//------------------------------------------------------------------------------
// SCADA FUXA : holding registers (FUXA 400001...), REAL = low word first (Float32MLE)
//------------------------------------------------------------------------------
	//--- DIP1500_1
	GVL_COM.COM_DIP1500_1.SCADA_INPUT_MOTOR_SPEED.Word_value[0]                                := GVL_MODBUS.Holding_register_TCP_HMI[0];    // 1 | DIP1500 Motor Speed (low word)
	GVL_COM.COM_DIP1500_1.SCADA_INPUT_MOTOR_SPEED.Word_value[1]                                := GVL_MODBUS.Holding_register_TCP_HMI[1];    // 2 | DIP1500 Motor Speed (high word)
	GVL_COM.COM_DIP1500_1.SCADA_INPUT_MAX_MOTOR_SPEED.Word_value[0]                            := GVL_MODBUS.Holding_register_TCP_HMI[2];    // 3 | DIP1500 Max Motor Speed (low word)
	GVL_COM.COM_DIP1500_1.SCADA_INPUT_MAX_MOTOR_SPEED.Word_value[1]                            := GVL_MODBUS.Holding_register_TCP_HMI[3];    // 4 | DIP1500 Max Motor Speed (high word)
	GVL_COM.COM_DIP1500_1.SCADA_INPUT_RUN_TIME_OR_VOLUME_SETPOINT.Word_value[0]                := GVL_MODBUS.Holding_register_TCP_HMI[4];    // 5 | DIP1500 Run Time Or Volume Setpoint (low word)
	GVL_COM.COM_DIP1500_1.SCADA_INPUT_RUN_TIME_OR_VOLUME_SETPOINT.Word_value[1]                := GVL_MODBUS.Holding_register_TCP_HMI[5];    // 6 | DIP1500 Run Time Or Volume Setpoint (high word)
	GVL_COM.COM_DIP1500_1.SCADA_INPUT_FLOW_RATE_OR_SPEED_CALIBRATION_COEFFICIENT.Word_value[0] := GVL_MODBUS.Holding_register_TCP_HMI[6];    // 7 | DIP1500 Flow Rate Or Speed Calibration Coefficient (low word)
	GVL_COM.COM_DIP1500_1.SCADA_INPUT_FLOW_RATE_OR_SPEED_CALIBRATION_COEFFICIENT.Word_value[1] := GVL_MODBUS.Holding_register_TCP_HMI[7];    // 8 | DIP1500 Flow Rate Or Speed Calibration Coefficient (high word)
	GVL_COM.COM_DIP1500_1.SCADA_INPUT_FOOT_SWITCH_INPUT_MODE                                   := GVL_MODBUS.Holding_register_TCP_HMI[8];    // 9 | DIP1500 Foot Switch Input Mode
	GVL_COM.COM_DIP1500_1.SCADA_INPUT_LIQUID_LEVEL_INPUT_MODE                                  := GVL_MODBUS.Holding_register_TCP_HMI[9];    // 10 | DIP1500 Liquid Level Input Mode
	GVL_COM.COM_DIP1500_1.SCADA_INPUT_STATE_OUTPUT_MODE                                        := GVL_MODBUS.Holding_register_TCP_HMI[10];   // 11 | DIP1500 State Output Mode
	GVL_COM.COM_DIP1500_1.SCADA_INPUT_COMMUNICATION_ADDRESS                                    := GVL_MODBUS.Holding_register_TCP_HMI[11];   // 12 | DIP1500 Communication Address
	GVL_COM.COM_DIP1500_1.SCADA_INPUT_BAUD_RATE_INDEX                                          := GVL_MODBUS.Holding_register_TCP_HMI[12];   // 13 | DIP1500 Baud Rate Index


//------------------------------------------------------------------------------
// HMI : coils (1001...)
//------------------------------------------------------------------------------
	//--- DOSENSOR_1
	GVL_COM.COM_DOSENSOR_1.HMI_INPUT_CALIBRATION_HIGH := GVL_MODBUS.Coils_TCP_HMI[125].0;   // 1001 | DO Calibration High
	GVL_COM.COM_DOSENSOR_1.HMI_INPUT_CALIBRATION_LOW  := GVL_MODBUS.Coils_TCP_HMI[125].1;   // 1002 | DO Calibration Low
	GVL_COM.COM_DOSENSOR_1.HMI_INPUT_LOCAL_REQUEST    := GVL_MODBUS.Coils_TCP_HMI[125].7;   // 1008 | DO Sensor Local Request
	GVL_COM.COM_DOSENSOR_1.HMI_INPUT_AUTO_REQUEST     := GVL_MODBUS.Coils_TCP_HMI[126].0;   // 1009 | DO Sensor Auto Request

	//--- DIP1500_1
	GVL_COM.COM_DIP1500_1.HMI_INPUT_MOTOR_START_STOP   := GVL_MODBUS.Coils_TCP_HMI[125].2;   // 1003 | DIP1500 Motor Start Stop
	GVL_COM.COM_DIP1500_1.HMI_INPUT_MOTOR_DIRECTION    := GVL_MODBUS.Coils_TCP_HMI[125].3;   // 1004 | DIP1500 Motor Direction
	GVL_COM.COM_DIP1500_1.HMI_INPUT_FLASH_SAVE         := GVL_MODBUS.Coils_TCP_HMI[125].4;   // 1005 | DIP1500 Flash Save
	GVL_COM.COM_DIP1500_1.HMI_INPUT_OPERATION_MODE     := GVL_MODBUS.Coils_TCP_HMI[125].5;   // 1006 | DIP1500 Operation Mode
	GVL_COM.COM_DIP1500_1.HMI_INPUT_PARAM_WRITE_ENABLE := GVL_MODBUS.Coils_TCP_HMI[125].6;   // 1007 | DIP1500 Parameter Write Enable
	GVL_COM.COM_DIP1500_1.HMI_INPUT_LOCAL_REQUEST      := GVL_MODBUS.Coils_TCP_HMI[126].1;   // 1010 | DIP1500 Local Request
	GVL_COM.COM_DIP1500_1.HMI_INPUT_AUTO_REQUEST       := GVL_MODBUS.Coils_TCP_HMI[126].2;   // 1011 | DIP1500 Auto Request

	//--- ADM100W_1
	GVL_COM.COM_ADM100W_1.HMI_INPUT_LOCAL_REQUEST := GVL_MODBUS.Coils_TCP_HMI[126].3;   // 1012 | ADM100W Local Request
	GVL_COM.COM_ADM100W_1.HMI_INPUT_AUTO_REQUEST  := GVL_MODBUS.Coils_TCP_HMI[126].4;   // 1013 | ADM100W Auto Request

	//--- UPI_LOCAL_HMI
	GVL_COM.COM_UPI_LOCAL_HMI.HMI_INPUT_LOCAL_REQUEST := GVL_MODBUS.Coils_TCP_HMI[126].5;   // 1014 | Global Local HMI Request
	GVL_COM.COM_UPI_LOCAL_HMI.HMI_INPUT_AUTO_REQUEST  := GVL_MODBUS.Coils_TCP_HMI[126].6;   // 1015 | Global Auto HMI Request


//------------------------------------------------------------------------------
// HMI : holding registers (1001...), REAL = low word first
//------------------------------------------------------------------------------
	//--- DIP1500_1
	GVL_COM.COM_DIP1500_1.HMI_INPUT_MOTOR_SPEED.Word_value[0]                                := GVL_MODBUS.Holding_register_TCP_HMI[1000];   // 1001 | DIP1500 Motor Speed (low word)
	GVL_COM.COM_DIP1500_1.HMI_INPUT_MOTOR_SPEED.Word_value[1]                                := GVL_MODBUS.Holding_register_TCP_HMI[1001];   // 1002 | DIP1500 Motor Speed (high word)
	GVL_COM.COM_DIP1500_1.HMI_INPUT_MAX_MOTOR_SPEED.Word_value[0]                            := GVL_MODBUS.Holding_register_TCP_HMI[1002];   // 1003 | DIP1500 Max Motor Speed (low word)
	GVL_COM.COM_DIP1500_1.HMI_INPUT_MAX_MOTOR_SPEED.Word_value[1]                            := GVL_MODBUS.Holding_register_TCP_HMI[1003];   // 1004 | DIP1500 Max Motor Speed (high word)
	GVL_COM.COM_DIP1500_1.HMI_INPUT_RUN_TIME_OR_VOLUME_SETPOINT.Word_value[0]                := GVL_MODBUS.Holding_register_TCP_HMI[1004];   // 1005 | DIP1500 Run Time Or Volume Setpoint (low word)
	GVL_COM.COM_DIP1500_1.HMI_INPUT_RUN_TIME_OR_VOLUME_SETPOINT.Word_value[1]                := GVL_MODBUS.Holding_register_TCP_HMI[1005];   // 1006 | DIP1500 Run Time Or Volume Setpoint (high word)
	GVL_COM.COM_DIP1500_1.HMI_INPUT_FLOW_RATE_OR_SPEED_CALIBRATION_COEFFICIENT.Word_value[0] := GVL_MODBUS.Holding_register_TCP_HMI[1006];   // 1007 | DIP1500 Flow Rate Or Speed Calibration Coefficient (low word)
	GVL_COM.COM_DIP1500_1.HMI_INPUT_FLOW_RATE_OR_SPEED_CALIBRATION_COEFFICIENT.Word_value[1] := GVL_MODBUS.Holding_register_TCP_HMI[1007];   // 1008 | DIP1500 Flow Rate Or Speed Calibration Coefficient (high word)
	GVL_COM.COM_DIP1500_1.HMI_INPUT_FOOT_SWITCH_INPUT_MODE                                   := GVL_MODBUS.Holding_register_TCP_HMI[1008];   // 1009 | DIP1500 Foot Switch Input Mode
	GVL_COM.COM_DIP1500_1.HMI_INPUT_LIQUID_LEVEL_INPUT_MODE                                  := GVL_MODBUS.Holding_register_TCP_HMI[1009];   // 1010 | DIP1500 Liquid Level Input Mode
	GVL_COM.COM_DIP1500_1.HMI_INPUT_STATE_OUTPUT_MODE                                        := GVL_MODBUS.Holding_register_TCP_HMI[1010];   // 1011 | DIP1500 State Output Mode
	GVL_COM.COM_DIP1500_1.HMI_INPUT_COMMUNICATION_ADDRESS                                    := GVL_MODBUS.Holding_register_TCP_HMI[1011];   // 1012 | DIP1500 Communication Address
	GVL_COM.COM_DIP1500_1.HMI_INPUT_BAUD_RATE_INDEX                                          := GVL_MODBUS.Holding_register_TCP_HMI[1012];   // 1013 | DIP1500 Baud Rate Index

GFC_COM_IN := TRUE;

                
END_FUNCTION

FUNCTION GFC_COM_OUT : BOOL

                  
//==============================================================================
// GFC_COM_OUT
// GVL_COM -> Modbus (GVL_MODBUS) : RTU equipment, SCADA FUXA, HMI
// Simple copies only, no conversion (conversions are done in the FBs)
//==============================================================================

//------------------------------------------------------------------------------
// COM : Modbus RTU, to equipment (write triggers are mapped directly in the slave I/O mapping)
//------------------------------------------------------------------------------
	//--- DIP1500_1
	GVL_MODBUS.DIP1500_Coils          := GVL_COM.COM_DIP1500_1.COM_OUTPUT_COILS;       // Coils 0x0001..0x0004
	GVL_MODBUS.DIP1500_Holding_Cmd    := GVL_COM.COM_DIP1500_1.COM_OUTPUT_HR_CMD;      // Holding registers 0x4001..0x4006
	GVL_MODBUS.DIP1500_Holding_Config := GVL_COM.COM_DIP1500_1.COM_OUTPUT_HR_CONFIG;   // Holding registers 0x400B..0x4011


//------------------------------------------------------------------------------
// SCADA FUXA : discrete inputs (FUXA 100001...)
//------------------------------------------------------------------------------
	//--- DOSENSOR_1
	GVL_MODBUS.Discret_input_TCP_HMI[0].0 := GVL_COM.COM_DOSENSOR_1.SCADA_OUTPUT_FAULT;               // 10001 | Do sensor fault
	GVL_MODBUS.Discret_input_TCP_HMI[0].1 := GVL_COM.COM_DOSENSOR_1.SCADA_OUTPUT_CALIBRATION_DONE;    // 10002 | Do sensor calibration done
	GVL_MODBUS.Discret_input_TCP_HMI[1].4 := GVL_COM.COM_DOSENSOR_1.SCADA_OUTPUT_LOCAL_FUXA_ACTIVE;   // 10013 | DO Sensor Local FUXA Active
	GVL_MODBUS.Discret_input_TCP_HMI[1].5 := GVL_COM.COM_DOSENSOR_1.SCADA_OUTPUT_LOCAL_HMI_ACTIVE;    // 10014 | DO Sensor Local HMI Active

	//--- ADM100W_1
	GVL_MODBUS.Discret_input_TCP_HMI[0].2 := GVL_COM.COM_ADM100W_1.SCADA_OUTPUT_ALARM_1_STATUS;      // 10003 | ADM100W Alarm 1 Status
	GVL_MODBUS.Discret_input_TCP_HMI[0].3 := GVL_COM.COM_ADM100W_1.SCADA_OUTPUT_ALARM_2_STATUS;      // 10004 | ADM100W Alarm 2 Status
	GVL_MODBUS.Discret_input_TCP_HMI[0].4 := GVL_COM.COM_ADM100W_1.SCADA_OUTPUT_ALARM_3_STATUS;      // 10005 | ADM100W Alarm 3 Status
	GVL_MODBUS.Discret_input_TCP_HMI[0].5 := GVL_COM.COM_ADM100W_1.SCADA_OUTPUT_ALARM_4_STATUS;      // 10006 | ADM100W Alarm 4 Status
	GVL_MODBUS.Discret_input_TCP_HMI[0].6 := GVL_COM.COM_ADM100W_1.SCADA_OUTPUT_ALARM_5_STATUS;      // 10007 | ADM100W Alarm 5 Status
	GVL_MODBUS.Discret_input_TCP_HMI[0].7 := GVL_COM.COM_ADM100W_1.SCADA_OUTPUT_ALARM_6_STATUS;      // 10008 | ADM100W Alarm 6 Status
	GVL_MODBUS.Discret_input_TCP_HMI[1].0 := GVL_COM.COM_ADM100W_1.SCADA_OUTPUT_ALARM_7_STATUS;      // 10009 | ADM100W Alarm 7 Status
	GVL_MODBUS.Discret_input_TCP_HMI[1].1 := GVL_COM.COM_ADM100W_1.SCADA_OUTPUT_ALARM_8_STATUS;      // 10010 | ADM100W Alarm 8 Status
	GVL_MODBUS.Discret_input_TCP_HMI[1].2 := GVL_COM.COM_ADM100W_1.SCADA_OUTPUT_ALARM_9_STATUS;      // 10011 | ADM100W Alarm 9 Status
	GVL_MODBUS.Discret_input_TCP_HMI[1].3 := GVL_COM.COM_ADM100W_1.SCADA_OUTPUT_ALARM_10_STATUS;     // 10012 | ADM100W Alarm 10 Status
	GVL_MODBUS.Discret_input_TCP_HMI[2].0 := GVL_COM.COM_ADM100W_1.SCADA_OUTPUT_LOCAL_FUXA_ACTIVE;   // 10017 | ADM100W Local FUXA Active
	GVL_MODBUS.Discret_input_TCP_HMI[2].1 := GVL_COM.COM_ADM100W_1.SCADA_OUTPUT_LOCAL_HMI_ACTIVE;    // 10018 | ADM100W Local HMI Active

	//--- DIP1500_1
	GVL_MODBUS.Discret_input_TCP_HMI[1].6 := GVL_COM.COM_DIP1500_1.SCADA_OUTPUT_LOCAL_FUXA_ACTIVE;   // 10015 | DIP1500 Local FUXA Active
	GVL_MODBUS.Discret_input_TCP_HMI[1].7 := GVL_COM.COM_DIP1500_1.SCADA_OUTPUT_LOCAL_HMI_ACTIVE;    // 10016 | DIP1500 Local HMI Active

	//--- UPI_LOCAL_FUXA
	GVL_MODBUS.Discret_input_TCP_HMI[2].2 := GVL_COM.COM_UPI_LOCAL_FUXA.SCADA_OUTPUT_LOCAL_ACTIVE;   // 10019 | Global Local FUXA Active

	//--- UPI_LOCAL_HMI
	GVL_MODBUS.Discret_input_TCP_HMI[2].3 := GVL_COM.COM_UPI_LOCAL_HMI.SCADA_OUTPUT_LOCAL_ACTIVE;   // 10020 | Global Local HMI Active


//------------------------------------------------------------------------------
// SCADA FUXA : input registers (FUXA 300001...), REAL = low word first (Float32MLE)
//------------------------------------------------------------------------------
	//--- ADM100W_1
	GVL_MODBUS.Input_register_TCP_HMI[0]  := GVL_COM.COM_ADM100W_1.SCADA_OUTPUT_FREQUENCY.Word_value[0];                   // 1 | ADM100W Frequency (low word)
	GVL_MODBUS.Input_register_TCP_HMI[1]  := GVL_COM.COM_ADM100W_1.SCADA_OUTPUT_FREQUENCY.Word_value[1];                   // 2 | ADM100W Frequency (high word)
	GVL_MODBUS.Input_register_TCP_HMI[2]  := GVL_COM.COM_ADM100W_1.SCADA_OUTPUT_L1_L2_VOLTAGE.Word_value[0];               // 3 | ADM100W L1-L2 Voltage (low word)
	GVL_MODBUS.Input_register_TCP_HMI[3]  := GVL_COM.COM_ADM100W_1.SCADA_OUTPUT_L1_L2_VOLTAGE.Word_value[1];               // 4 | ADM100W L1-L2 Voltage (high word)
	GVL_MODBUS.Input_register_TCP_HMI[4]  := GVL_COM.COM_ADM100W_1.SCADA_OUTPUT_L1_N_VOLTAGE.Word_value[0];                // 5 | ADM100W L1-N Voltage (low word)
	GVL_MODBUS.Input_register_TCP_HMI[5]  := GVL_COM.COM_ADM100W_1.SCADA_OUTPUT_L1_N_VOLTAGE.Word_value[1];                // 6 | ADM100W L1-N Voltage (high word)
	GVL_MODBUS.Input_register_TCP_HMI[6]  := GVL_COM.COM_ADM100W_1.SCADA_OUTPUT_L1_CURRENT.Word_value[0];                  // 7 | ADM100W L1 Current (low word)
	GVL_MODBUS.Input_register_TCP_HMI[7]  := GVL_COM.COM_ADM100W_1.SCADA_OUTPUT_L1_CURRENT.Word_value[1];                  // 8 | ADM100W L1 Current (high word)
	GVL_MODBUS.Input_register_TCP_HMI[8]  := GVL_COM.COM_ADM100W_1.SCADA_OUTPUT_L1_ACTIVE_POWER.Word_value[0];             // 9 | ADM100W L1 Active Power (low word)
	GVL_MODBUS.Input_register_TCP_HMI[9]  := GVL_COM.COM_ADM100W_1.SCADA_OUTPUT_L1_ACTIVE_POWER.Word_value[1];             // 10 | ADM100W L1 Active Power (high word)
	GVL_MODBUS.Input_register_TCP_HMI[10] := GVL_COM.COM_ADM100W_1.SCADA_OUTPUT_L1_APPARENT_POWER.Word_value[0];           // 11 | ADM100W L1 Apparent Power (low word)
	GVL_MODBUS.Input_register_TCP_HMI[11] := GVL_COM.COM_ADM100W_1.SCADA_OUTPUT_L1_APPARENT_POWER.Word_value[1];           // 12 | ADM100W L1 Apparent Power (high word)
	GVL_MODBUS.Input_register_TCP_HMI[12] := GVL_COM.COM_ADM100W_1.SCADA_OUTPUT_L1_REACTIVE_POWER.Word_value[0];           // 13 | ADM100W L1 Reactive Power (low word)
	GVL_MODBUS.Input_register_TCP_HMI[13] := GVL_COM.COM_ADM100W_1.SCADA_OUTPUT_L1_REACTIVE_POWER.Word_value[1];           // 14 | ADM100W L1 Reactive Power (high word)
	GVL_MODBUS.Input_register_TCP_HMI[14] := GVL_COM.COM_ADM100W_1.SCADA_OUTPUT_L1_CURRENT_PHASE_ANGLE.Word_value[0];      // 15 | ADM100W L1 Current Phase Angle (low word)
	GVL_MODBUS.Input_register_TCP_HMI[15] := GVL_COM.COM_ADM100W_1.SCADA_OUTPUT_L1_CURRENT_PHASE_ANGLE.Word_value[1];      // 16 | ADM100W L1 Current Phase Angle (high word)
	GVL_MODBUS.Input_register_TCP_HMI[16] := GVL_COM.COM_ADM100W_1.SCADA_OUTPUT_L1_POWER_FACTOR.Word_value[0];             // 17 | ADM100W L1 Power Factor (low word)
	GVL_MODBUS.Input_register_TCP_HMI[17] := GVL_COM.COM_ADM100W_1.SCADA_OUTPUT_L1_POWER_FACTOR.Word_value[1];             // 18 | ADM100W L1 Power Factor (high word)
	GVL_MODBUS.Input_register_TCP_HMI[18] := GVL_COM.COM_ADM100W_1.SCADA_OUTPUT_L1_VOLTAGE_THD.Word_value[0];              // 19 | ADM100W L1 Voltage THD (low word)
	GVL_MODBUS.Input_register_TCP_HMI[19] := GVL_COM.COM_ADM100W_1.SCADA_OUTPUT_L1_VOLTAGE_THD.Word_value[1];              // 20 | ADM100W L1 Voltage THD (high word)
	GVL_MODBUS.Input_register_TCP_HMI[20] := GVL_COM.COM_ADM100W_1.SCADA_OUTPUT_L1_CURRENT_THD.Word_value[0];              // 21 | ADM100W L1 Current THD (low word)
	GVL_MODBUS.Input_register_TCP_HMI[21] := GVL_COM.COM_ADM100W_1.SCADA_OUTPUT_L1_CURRENT_THD.Word_value[1];              // 22 | ADM100W L1 Current THD (high word)
	GVL_MODBUS.Input_register_TCP_HMI[22] := GVL_COM.COM_ADM100W_1.SCADA_OUTPUT_L1_MAX_LOAD.Word_value[0];                 // 23 | ADM100W L1 Max Load (low word)
	GVL_MODBUS.Input_register_TCP_HMI[23] := GVL_COM.COM_ADM100W_1.SCADA_OUTPUT_L1_MAX_LOAD.Word_value[1];                 // 24 | ADM100W L1 Max Load (high word)
	GVL_MODBUS.Input_register_TCP_HMI[24] := GVL_COM.COM_ADM100W_1.SCADA_OUTPUT_L1_L2_VOLTAGE_PHASE_ANGLE.Word_value[0];   // 25 | ADM100W L1-L2 Voltage Phase Angle (low word)
	GVL_MODBUS.Input_register_TCP_HMI[25] := GVL_COM.COM_ADM100W_1.SCADA_OUTPUT_L1_L2_VOLTAGE_PHASE_ANGLE.Word_value[1];   // 26 | ADM100W L1-L2 Voltage Phase Angle (high word)
	GVL_MODBUS.Input_register_TCP_HMI[26] := GVL_COM.COM_ADM100W_1.SCADA_OUTPUT_L2_L3_VOLTAGE.Word_value[0];               // 27 | ADM100W L2-L3 Voltage (low word)
	GVL_MODBUS.Input_register_TCP_HMI[27] := GVL_COM.COM_ADM100W_1.SCADA_OUTPUT_L2_L3_VOLTAGE.Word_value[1];               // 28 | ADM100W L2-L3 Voltage (high word)
	GVL_MODBUS.Input_register_TCP_HMI[28] := GVL_COM.COM_ADM100W_1.SCADA_OUTPUT_L2_N_VOLTAGE.Word_value[0];                // 29 | ADM100W L2-N Voltage (low word)
	GVL_MODBUS.Input_register_TCP_HMI[29] := GVL_COM.COM_ADM100W_1.SCADA_OUTPUT_L2_N_VOLTAGE.Word_value[1];                // 30 | ADM100W L2-N Voltage (high word)
	GVL_MODBUS.Input_register_TCP_HMI[30] := GVL_COM.COM_ADM100W_1.SCADA_OUTPUT_L2_CURRENT.Word_value[0];                  // 31 | ADM100W L2 Current (low word)
	GVL_MODBUS.Input_register_TCP_HMI[31] := GVL_COM.COM_ADM100W_1.SCADA_OUTPUT_L2_CURRENT.Word_value[1];                  // 32 | ADM100W L2 Current (high word)
	GVL_MODBUS.Input_register_TCP_HMI[32] := GVL_COM.COM_ADM100W_1.SCADA_OUTPUT_L2_ACTIVE_POWER.Word_value[0];             // 33 | ADM100W L2 Active Power (low word)
	GVL_MODBUS.Input_register_TCP_HMI[33] := GVL_COM.COM_ADM100W_1.SCADA_OUTPUT_L2_ACTIVE_POWER.Word_value[1];             // 34 | ADM100W L2 Active Power (high word)
	GVL_MODBUS.Input_register_TCP_HMI[34] := GVL_COM.COM_ADM100W_1.SCADA_OUTPUT_L2_APPARENT_POWER.Word_value[0];           // 35 | ADM100W L2 Apparent Power (low word)
	GVL_MODBUS.Input_register_TCP_HMI[35] := GVL_COM.COM_ADM100W_1.SCADA_OUTPUT_L2_APPARENT_POWER.Word_value[1];           // 36 | ADM100W L2 Apparent Power (high word)
	GVL_MODBUS.Input_register_TCP_HMI[36] := GVL_COM.COM_ADM100W_1.SCADA_OUTPUT_L2_REACTIVE_POWER.Word_value[0];           // 37 | ADM100W L2 Reactive Power (low word)
	GVL_MODBUS.Input_register_TCP_HMI[37] := GVL_COM.COM_ADM100W_1.SCADA_OUTPUT_L2_REACTIVE_POWER.Word_value[1];           // 38 | ADM100W L2 Reactive Power (high word)
	GVL_MODBUS.Input_register_TCP_HMI[38] := GVL_COM.COM_ADM100W_1.SCADA_OUTPUT_L2_CURRENT_PHASE_ANGLE.Word_value[0];      // 39 | ADM100W L2 Current Phase Angle (low word)
	GVL_MODBUS.Input_register_TCP_HMI[39] := GVL_COM.COM_ADM100W_1.SCADA_OUTPUT_L2_CURRENT_PHASE_ANGLE.Word_value[1];      // 40 | ADM100W L2 Current Phase Angle (high word)
	GVL_MODBUS.Input_register_TCP_HMI[40] := GVL_COM.COM_ADM100W_1.SCADA_OUTPUT_L2_POWER_FACTOR.Word_value[0];             // 41 | ADM100W L2 Power Factor (low word)
	GVL_MODBUS.Input_register_TCP_HMI[41] := GVL_COM.COM_ADM100W_1.SCADA_OUTPUT_L2_POWER_FACTOR.Word_value[1];             // 42 | ADM100W L2 Power Factor (high word)
	GVL_MODBUS.Input_register_TCP_HMI[42] := GVL_COM.COM_ADM100W_1.SCADA_OUTPUT_L2_VOLTAGE_THD.Word_value[0];              // 43 | ADM100W L2 Voltage THD (low word)
	GVL_MODBUS.Input_register_TCP_HMI[43] := GVL_COM.COM_ADM100W_1.SCADA_OUTPUT_L2_VOLTAGE_THD.Word_value[1];              // 44 | ADM100W L2 Voltage THD (high word)
	GVL_MODBUS.Input_register_TCP_HMI[44] := GVL_COM.COM_ADM100W_1.SCADA_OUTPUT_L2_CURRENT_THD.Word_value[0];              // 45 | ADM100W L2 Current THD (low word)
	GVL_MODBUS.Input_register_TCP_HMI[45] := GVL_COM.COM_ADM100W_1.SCADA_OUTPUT_L2_CURRENT_THD.Word_value[1];              // 46 | ADM100W L2 Current THD (high word)
	GVL_MODBUS.Input_register_TCP_HMI[46] := GVL_COM.COM_ADM100W_1.SCADA_OUTPUT_L2_MAX_LOAD.Word_value[0];                 // 47 | ADM100W L2 Max Load (low word)
	GVL_MODBUS.Input_register_TCP_HMI[47] := GVL_COM.COM_ADM100W_1.SCADA_OUTPUT_L2_MAX_LOAD.Word_value[1];                 // 48 | ADM100W L2 Max Load (high word)
	GVL_MODBUS.Input_register_TCP_HMI[48] := GVL_COM.COM_ADM100W_1.SCADA_OUTPUT_L1_L3_VOLTAGE_PHASE_ANGLE.Word_value[0];   // 49 | ADM100W L1-L3 Voltage Phase Angle (low word)
	GVL_MODBUS.Input_register_TCP_HMI[49] := GVL_COM.COM_ADM100W_1.SCADA_OUTPUT_L1_L3_VOLTAGE_PHASE_ANGLE.Word_value[1];   // 50 | ADM100W L1-L3 Voltage Phase Angle (high word)
	GVL_MODBUS.Input_register_TCP_HMI[50] := GVL_COM.COM_ADM100W_1.SCADA_OUTPUT_L3_L1_VOLTAGE.Word_value[0];               // 51 | ADM100W L3-L1 Voltage (low word)
	GVL_MODBUS.Input_register_TCP_HMI[51] := GVL_COM.COM_ADM100W_1.SCADA_OUTPUT_L3_L1_VOLTAGE.Word_value[1];               // 52 | ADM100W L3-L1 Voltage (high word)
	GVL_MODBUS.Input_register_TCP_HMI[52] := GVL_COM.COM_ADM100W_1.SCADA_OUTPUT_L3_N_VOLTAGE.Word_value[0];                // 53 | ADM100W L3-N Voltage (low word)
	GVL_MODBUS.Input_register_TCP_HMI[53] := GVL_COM.COM_ADM100W_1.SCADA_OUTPUT_L3_N_VOLTAGE.Word_value[1];                // 54 | ADM100W L3-N Voltage (high word)
	GVL_MODBUS.Input_register_TCP_HMI[54] := GVL_COM.COM_ADM100W_1.SCADA_OUTPUT_L3_CURRENT.Word_value[0];                  // 55 | ADM100W L3 Current (low word)
	GVL_MODBUS.Input_register_TCP_HMI[55] := GVL_COM.COM_ADM100W_1.SCADA_OUTPUT_L3_CURRENT.Word_value[1];                  // 56 | ADM100W L3 Current (high word)
	GVL_MODBUS.Input_register_TCP_HMI[56] := GVL_COM.COM_ADM100W_1.SCADA_OUTPUT_L3_ACTIVE_POWER.Word_value[0];             // 57 | ADM100W L3 Active Power (low word)
	GVL_MODBUS.Input_register_TCP_HMI[57] := GVL_COM.COM_ADM100W_1.SCADA_OUTPUT_L3_ACTIVE_POWER.Word_value[1];             // 58 | ADM100W L3 Active Power (high word)
	GVL_MODBUS.Input_register_TCP_HMI[58] := GVL_COM.COM_ADM100W_1.SCADA_OUTPUT_L3_APPARENT_POWER.Word_value[0];           // 59 | ADM100W L3 Apparent Power (low word)
	GVL_MODBUS.Input_register_TCP_HMI[59] := GVL_COM.COM_ADM100W_1.SCADA_OUTPUT_L3_APPARENT_POWER.Word_value[1];           // 60 | ADM100W L3 Apparent Power (high word)
	GVL_MODBUS.Input_register_TCP_HMI[60] := GVL_COM.COM_ADM100W_1.SCADA_OUTPUT_L3_REACTIVE_POWER.Word_value[0];           // 61 | ADM100W L3 Reactive Power (low word)
	GVL_MODBUS.Input_register_TCP_HMI[61] := GVL_COM.COM_ADM100W_1.SCADA_OUTPUT_L3_REACTIVE_POWER.Word_value[1];           // 62 | ADM100W L3 Reactive Power (high word)
	GVL_MODBUS.Input_register_TCP_HMI[62] := GVL_COM.COM_ADM100W_1.SCADA_OUTPUT_L3_CURRENT_PHASE_ANGLE.Word_value[0];      // 63 | ADM100W L3 Current Phase Angle (low word)
	GVL_MODBUS.Input_register_TCP_HMI[63] := GVL_COM.COM_ADM100W_1.SCADA_OUTPUT_L3_CURRENT_PHASE_ANGLE.Word_value[1];      // 64 | ADM100W L3 Current Phase Angle (high word)
	GVL_MODBUS.Input_register_TCP_HMI[64] := GVL_COM.COM_ADM100W_1.SCADA_OUTPUT_L3_POWER_FACTOR.Word_value[0];             // 65 | ADM100W L3 Power Factor (low word)
	GVL_MODBUS.Input_register_TCP_HMI[65] := GVL_COM.COM_ADM100W_1.SCADA_OUTPUT_L3_POWER_FACTOR.Word_value[1];             // 66 | ADM100W L3 Power Factor (high word)
	GVL_MODBUS.Input_register_TCP_HMI[66] := GVL_COM.COM_ADM100W_1.SCADA_OUTPUT_L3_VOLTAGE_THD.Word_value[0];              // 67 | ADM100W L3 Voltage THD (low word)
	GVL_MODBUS.Input_register_TCP_HMI[67] := GVL_COM.COM_ADM100W_1.SCADA_OUTPUT_L3_VOLTAGE_THD.Word_value[1];              // 68 | ADM100W L3 Voltage THD (high word)
	GVL_MODBUS.Input_register_TCP_HMI[68] := GVL_COM.COM_ADM100W_1.SCADA_OUTPUT_L3_CURRENT_THD.Word_value[0];              // 69 | ADM100W L3 Current THD (low word)
	GVL_MODBUS.Input_register_TCP_HMI[69] := GVL_COM.COM_ADM100W_1.SCADA_OUTPUT_L3_CURRENT_THD.Word_value[1];              // 70 | ADM100W L3 Current THD (high word)
	GVL_MODBUS.Input_register_TCP_HMI[70] := GVL_COM.COM_ADM100W_1.SCADA_OUTPUT_L3_MAX_LOAD.Word_value[0];                 // 71 | ADM100W L3 Max Load (low word)
	GVL_MODBUS.Input_register_TCP_HMI[71] := GVL_COM.COM_ADM100W_1.SCADA_OUTPUT_L3_MAX_LOAD.Word_value[1];                 // 72 | ADM100W L3 Max Load (high word)
	GVL_MODBUS.Input_register_TCP_HMI[72] := GVL_COM.COM_ADM100W_1.SCADA_OUTPUT_INTERNAL_TEMPERATURE.Word_value[0];        // 73 | ADM100W Internal Temperature (low word)
	GVL_MODBUS.Input_register_TCP_HMI[73] := GVL_COM.COM_ADM100W_1.SCADA_OUTPUT_INTERNAL_TEMPERATURE.Word_value[1];        // 74 | ADM100W Internal Temperature (high word)
	GVL_MODBUS.Input_register_TCP_HMI[74] := GVL_COM.COM_ADM100W_1.SCADA_OUTPUT_ACTIVE_ENERGY.Word_value[0];               // 75 | ADM100W Active Energy (low word)
	GVL_MODBUS.Input_register_TCP_HMI[75] := GVL_COM.COM_ADM100W_1.SCADA_OUTPUT_ACTIVE_ENERGY.Word_value[1];               // 76 | ADM100W Active Energy (high word)
	GVL_MODBUS.Input_register_TCP_HMI[76] := GVL_COM.COM_ADM100W_1.SCADA_OUTPUT_APPARENT_ENERGY.Word_value[0];             // 77 | ADM100W Apparent Energy (low word)
	GVL_MODBUS.Input_register_TCP_HMI[77] := GVL_COM.COM_ADM100W_1.SCADA_OUTPUT_APPARENT_ENERGY.Word_value[1];             // 78 | ADM100W Apparent Energy (high word)
	GVL_MODBUS.Input_register_TCP_HMI[78] := GVL_COM.COM_ADM100W_1.SCADA_OUTPUT_REACTIVE_ENERGY.Word_value[0];             // 79 | ADM100W Reactive Energy (low word)
	GVL_MODBUS.Input_register_TCP_HMI[79] := GVL_COM.COM_ADM100W_1.SCADA_OUTPUT_REACTIVE_ENERGY.Word_value[1];             // 80 | ADM100W Reactive Energy (high word)
	GVL_MODBUS.Input_register_TCP_HMI[80] := GVL_COM.COM_ADM100W_1.SCADA_OUTPUT_TOTAL_ACTIVE_POWER.Word_value[0];          // 81 | ADM100W Total Active Power (low word)
	GVL_MODBUS.Input_register_TCP_HMI[81] := GVL_COM.COM_ADM100W_1.SCADA_OUTPUT_TOTAL_ACTIVE_POWER.Word_value[1];          // 82 | ADM100W Total Active Power (high word)
	GVL_MODBUS.Input_register_TCP_HMI[82] := GVL_COM.COM_ADM100W_1.SCADA_OUTPUT_TOTAL_APPARENT_POWER.Word_value[0];        // 83 | ADM100W Total Apparent Power (low word)
	GVL_MODBUS.Input_register_TCP_HMI[83] := GVL_COM.COM_ADM100W_1.SCADA_OUTPUT_TOTAL_APPARENT_POWER.Word_value[1];        // 84 | ADM100W Total Apparent Power (high word)
	GVL_MODBUS.Input_register_TCP_HMI[84] := GVL_COM.COM_ADM100W_1.SCADA_OUTPUT_TOTAL_REACTIVE_POWER.Word_value[0];        // 85 | ADM100W Total Reactive Power (low word)
	GVL_MODBUS.Input_register_TCP_HMI[85] := GVL_COM.COM_ADM100W_1.SCADA_OUTPUT_TOTAL_REACTIVE_POWER.Word_value[1];        // 86 | ADM100W Total Reactive Power (high word)
	GVL_MODBUS.Input_register_TCP_HMI[86] := GVL_COM.COM_ADM100W_1.SCADA_OUTPUT_ALL_PHASE_POWER_FACTOR.Word_value[0];      // 87 | ADM100W All Phase Power Factor (low word)
	GVL_MODBUS.Input_register_TCP_HMI[87] := GVL_COM.COM_ADM100W_1.SCADA_OUTPUT_ALL_PHASE_POWER_FACTOR.Word_value[1];      // 88 | ADM100W All Phase Power Factor (high word)

	//--- DOSENSOR_1
	GVL_MODBUS.Input_register_TCP_HMI[88] := GVL_COM.COM_DOSENSOR_1.SCADA_OUTPUT_SIGNAL.Word_value[0];   // 89 | DO Sensor Signal (low word)
	GVL_MODBUS.Input_register_TCP_HMI[89] := GVL_COM.COM_DOSENSOR_1.SCADA_OUTPUT_SIGNAL.Word_value[1];   // 90 | DO Sensor Signal (high word)

	//--- DIP1500_1
	GVL_MODBUS.Input_register_TCP_HMI[90] := GVL_COM.COM_DIP1500_1.SCADA_OUTPUT_FIRMWARE_VERSION;                               // 91 | DIP1500 Firmware Version
	GVL_MODBUS.Input_register_TCP_HMI[91] := GVL_COM.COM_DIP1500_1.SCADA_OUTPUT_HARDWARE_VERSION;                               // 92 | DIP1500 Hardware Version
	GVL_MODBUS.Input_register_TCP_HMI[92] := GVL_COM.COM_DIP1500_1.SCADA_OUTPUT_TEMPERATURE;                                    // 93 | DIP1500 Temperature
	GVL_MODBUS.Input_register_TCP_HMI[93] := GVL_COM.COM_DIP1500_1.SCADA_OUTPUT_FLOAT_LEVEL_ALARM;                              // 94 | DIP1500 Float Level Alarm
	GVL_MODBUS.Input_register_TCP_HMI[94] := GVL_COM.COM_DIP1500_1.SCADA_OUTPUT_DIGITAL_OUTPUT_VALUE;                           // 95 | DIP1500 Digital Output Value
	GVL_MODBUS.Input_register_TCP_HMI[95] := GVL_COM.COM_DIP1500_1.SCADA_OUTPUT_REAL_TIME_RUN_TIME_OR_VOLUME.Word_value[0];     // 96 | DIP1500 Real-Time Run Time Or Volume (low word)
	GVL_MODBUS.Input_register_TCP_HMI[96] := GVL_COM.COM_DIP1500_1.SCADA_OUTPUT_REAL_TIME_RUN_TIME_OR_VOLUME.Word_value[1];     // 97 | DIP1500 Real-Time Run Time Or Volume (high word)
	GVL_MODBUS.Input_register_TCP_HMI[97] := GVL_COM.COM_DIP1500_1.SCADA_OUTPUT_ACCUMULATED_RUN_TIME_OR_VOLUME.Word_value[0];   // 98 | DIP1500 Accumulated Run Time Or Volume (low word)
	GVL_MODBUS.Input_register_TCP_HMI[98] := GVL_COM.COM_DIP1500_1.SCADA_OUTPUT_ACCUMULATED_RUN_TIME_OR_VOLUME.Word_value[1];   // 99 | DIP1500 Accumulated Run Time Or Volume (high word)


//------------------------------------------------------------------------------
// HMI : discrete inputs (11001...)
//------------------------------------------------------------------------------
	//--- DOSENSOR_1
	GVL_MODBUS.Discret_input_TCP_HMI[125].0 := GVL_COM.COM_DOSENSOR_1.HMI_OUTPUT_FAULT;              // 11001 | Do sensor fault
	GVL_MODBUS.Discret_input_TCP_HMI[125].1 := GVL_COM.COM_DOSENSOR_1.HMI_OUTPUT_CALIBRATION_DONE;   // 11002 | Do sensor calibration done
	GVL_MODBUS.Discret_input_TCP_HMI[126].5 := GVL_COM.COM_DOSENSOR_1.HMI_OUTPUT_LOCAL_ACTIVE;       // 11014 | DO Sensor Local Active

	//--- ADM100W_1
	GVL_MODBUS.Discret_input_TCP_HMI[125].2 := GVL_COM.COM_ADM100W_1.HMI_OUTPUT_ALARM_1_STATUS;    // 11003 | ADM100W Alarm 1 Status
	GVL_MODBUS.Discret_input_TCP_HMI[125].3 := GVL_COM.COM_ADM100W_1.HMI_OUTPUT_ALARM_2_STATUS;    // 11004 | ADM100W Alarm 2 Status
	GVL_MODBUS.Discret_input_TCP_HMI[125].4 := GVL_COM.COM_ADM100W_1.HMI_OUTPUT_ALARM_3_STATUS;    // 11005 | ADM100W Alarm 3 Status
	GVL_MODBUS.Discret_input_TCP_HMI[125].5 := GVL_COM.COM_ADM100W_1.HMI_OUTPUT_ALARM_4_STATUS;    // 11006 | ADM100W Alarm 4 Status
	GVL_MODBUS.Discret_input_TCP_HMI[125].6 := GVL_COM.COM_ADM100W_1.HMI_OUTPUT_ALARM_5_STATUS;    // 11007 | ADM100W Alarm 5 Status
	GVL_MODBUS.Discret_input_TCP_HMI[125].7 := GVL_COM.COM_ADM100W_1.HMI_OUTPUT_ALARM_6_STATUS;    // 11008 | ADM100W Alarm 6 Status
	GVL_MODBUS.Discret_input_TCP_HMI[126].0 := GVL_COM.COM_ADM100W_1.HMI_OUTPUT_ALARM_7_STATUS;    // 11009 | ADM100W Alarm 7 Status
	GVL_MODBUS.Discret_input_TCP_HMI[126].1 := GVL_COM.COM_ADM100W_1.HMI_OUTPUT_ALARM_8_STATUS;    // 11010 | ADM100W Alarm 8 Status
	GVL_MODBUS.Discret_input_TCP_HMI[126].2 := GVL_COM.COM_ADM100W_1.HMI_OUTPUT_ALARM_9_STATUS;    // 11011 | ADM100W Alarm 9 Status
	GVL_MODBUS.Discret_input_TCP_HMI[126].3 := GVL_COM.COM_ADM100W_1.HMI_OUTPUT_ALARM_10_STATUS;   // 11012 | ADM100W Alarm 10 Status
	GVL_MODBUS.Discret_input_TCP_HMI[127].1 := GVL_COM.COM_ADM100W_1.HMI_OUTPUT_LOCAL_ACTIVE;      // 11018 | ADM100W Local Active

	//--- DIP1500_1
	GVL_MODBUS.Discret_input_TCP_HMI[126].7 := GVL_COM.COM_DIP1500_1.HMI_OUTPUT_LOCAL_ACTIVE;   // 11016 | DIP1500 Local Active

	//--- UPI_LOCAL_HMI
	GVL_MODBUS.Discret_input_TCP_HMI[127].3 := GVL_COM.COM_UPI_LOCAL_HMI.HMI_OUTPUT_LOCAL_ACTIVE;   // 11020 | Global Local HMI Active


//------------------------------------------------------------------------------
// HMI : input registers (1001...), REAL = low word first
//------------------------------------------------------------------------------
	//--- ADM100W_1
	GVL_MODBUS.Input_register_TCP_HMI[1000] := GVL_COM.COM_ADM100W_1.HMI_OUTPUT_FREQUENCY.Word_value[0];                   // 1001 | ADM100W Frequency (low word)
	GVL_MODBUS.Input_register_TCP_HMI[1001] := GVL_COM.COM_ADM100W_1.HMI_OUTPUT_FREQUENCY.Word_value[1];                   // 1002 | ADM100W Frequency (high word)
	GVL_MODBUS.Input_register_TCP_HMI[1002] := GVL_COM.COM_ADM100W_1.HMI_OUTPUT_L1_L2_VOLTAGE.Word_value[0];               // 1003 | ADM100W L1-L2 Voltage (low word)
	GVL_MODBUS.Input_register_TCP_HMI[1003] := GVL_COM.COM_ADM100W_1.HMI_OUTPUT_L1_L2_VOLTAGE.Word_value[1];               // 1004 | ADM100W L1-L2 Voltage (high word)
	GVL_MODBUS.Input_register_TCP_HMI[1004] := GVL_COM.COM_ADM100W_1.HMI_OUTPUT_L1_N_VOLTAGE.Word_value[0];                // 1005 | ADM100W L1-N Voltage (low word)
	GVL_MODBUS.Input_register_TCP_HMI[1005] := GVL_COM.COM_ADM100W_1.HMI_OUTPUT_L1_N_VOLTAGE.Word_value[1];                // 1006 | ADM100W L1-N Voltage (high word)
	GVL_MODBUS.Input_register_TCP_HMI[1006] := GVL_COM.COM_ADM100W_1.HMI_OUTPUT_L1_CURRENT.Word_value[0];                  // 1007 | ADM100W L1 Current (low word)
	GVL_MODBUS.Input_register_TCP_HMI[1007] := GVL_COM.COM_ADM100W_1.HMI_OUTPUT_L1_CURRENT.Word_value[1];                  // 1008 | ADM100W L1 Current (high word)
	GVL_MODBUS.Input_register_TCP_HMI[1008] := GVL_COM.COM_ADM100W_1.HMI_OUTPUT_L1_ACTIVE_POWER.Word_value[0];             // 1009 | ADM100W L1 Active Power (low word)
	GVL_MODBUS.Input_register_TCP_HMI[1009] := GVL_COM.COM_ADM100W_1.HMI_OUTPUT_L1_ACTIVE_POWER.Word_value[1];             // 1010 | ADM100W L1 Active Power (high word)
	GVL_MODBUS.Input_register_TCP_HMI[1010] := GVL_COM.COM_ADM100W_1.HMI_OUTPUT_L1_APPARENT_POWER.Word_value[0];           // 1011 | ADM100W L1 Apparent Power (low word)
	GVL_MODBUS.Input_register_TCP_HMI[1011] := GVL_COM.COM_ADM100W_1.HMI_OUTPUT_L1_APPARENT_POWER.Word_value[1];           // 1012 | ADM100W L1 Apparent Power (high word)
	GVL_MODBUS.Input_register_TCP_HMI[1012] := GVL_COM.COM_ADM100W_1.HMI_OUTPUT_L1_REACTIVE_POWER.Word_value[0];           // 1013 | ADM100W L1 Reactive Power (low word)
	GVL_MODBUS.Input_register_TCP_HMI[1013] := GVL_COM.COM_ADM100W_1.HMI_OUTPUT_L1_REACTIVE_POWER.Word_value[1];           // 1014 | ADM100W L1 Reactive Power (high word)
	GVL_MODBUS.Input_register_TCP_HMI[1014] := GVL_COM.COM_ADM100W_1.HMI_OUTPUT_L1_CURRENT_PHASE_ANGLE.Word_value[0];      // 1015 | ADM100W L1 Current Phase Angle (low word)
	GVL_MODBUS.Input_register_TCP_HMI[1015] := GVL_COM.COM_ADM100W_1.HMI_OUTPUT_L1_CURRENT_PHASE_ANGLE.Word_value[1];      // 1016 | ADM100W L1 Current Phase Angle (high word)
	GVL_MODBUS.Input_register_TCP_HMI[1016] := GVL_COM.COM_ADM100W_1.HMI_OUTPUT_L1_POWER_FACTOR.Word_value[0];             // 1017 | ADM100W L1 Power Factor (low word)
	GVL_MODBUS.Input_register_TCP_HMI[1017] := GVL_COM.COM_ADM100W_1.HMI_OUTPUT_L1_POWER_FACTOR.Word_value[1];             // 1018 | ADM100W L1 Power Factor (high word)
	GVL_MODBUS.Input_register_TCP_HMI[1018] := GVL_COM.COM_ADM100W_1.HMI_OUTPUT_L1_VOLTAGE_THD.Word_value[0];              // 1019 | ADM100W L1 Voltage THD (low word)
	GVL_MODBUS.Input_register_TCP_HMI[1019] := GVL_COM.COM_ADM100W_1.HMI_OUTPUT_L1_VOLTAGE_THD.Word_value[1];              // 1020 | ADM100W L1 Voltage THD (high word)
	GVL_MODBUS.Input_register_TCP_HMI[1020] := GVL_COM.COM_ADM100W_1.HMI_OUTPUT_L1_CURRENT_THD.Word_value[0];              // 1021 | ADM100W L1 Current THD (low word)
	GVL_MODBUS.Input_register_TCP_HMI[1021] := GVL_COM.COM_ADM100W_1.HMI_OUTPUT_L1_CURRENT_THD.Word_value[1];              // 1022 | ADM100W L1 Current THD (high word)
	GVL_MODBUS.Input_register_TCP_HMI[1022] := GVL_COM.COM_ADM100W_1.HMI_OUTPUT_L1_MAX_LOAD.Word_value[0];                 // 1023 | ADM100W L1 Max Load (low word)
	GVL_MODBUS.Input_register_TCP_HMI[1023] := GVL_COM.COM_ADM100W_1.HMI_OUTPUT_L1_MAX_LOAD.Word_value[1];                 // 1024 | ADM100W L1 Max Load (high word)
	GVL_MODBUS.Input_register_TCP_HMI[1024] := GVL_COM.COM_ADM100W_1.HMI_OUTPUT_L1_L2_VOLTAGE_PHASE_ANGLE.Word_value[0];   // 1025 | ADM100W L1-L2 Voltage Phase Angle (low word)
	GVL_MODBUS.Input_register_TCP_HMI[1025] := GVL_COM.COM_ADM100W_1.HMI_OUTPUT_L1_L2_VOLTAGE_PHASE_ANGLE.Word_value[1];   // 1026 | ADM100W L1-L2 Voltage Phase Angle (high word)
	GVL_MODBUS.Input_register_TCP_HMI[1026] := GVL_COM.COM_ADM100W_1.HMI_OUTPUT_L2_L3_VOLTAGE.Word_value[0];               // 1027 | ADM100W L2-L3 Voltage (low word)
	GVL_MODBUS.Input_register_TCP_HMI[1027] := GVL_COM.COM_ADM100W_1.HMI_OUTPUT_L2_L3_VOLTAGE.Word_value[1];               // 1028 | ADM100W L2-L3 Voltage (high word)
	GVL_MODBUS.Input_register_TCP_HMI[1028] := GVL_COM.COM_ADM100W_1.HMI_OUTPUT_L2_N_VOLTAGE.Word_value[0];                // 1029 | ADM100W L2-N Voltage (low word)
	GVL_MODBUS.Input_register_TCP_HMI[1029] := GVL_COM.COM_ADM100W_1.HMI_OUTPUT_L2_N_VOLTAGE.Word_value[1];                // 1030 | ADM100W L2-N Voltage (high word)
	GVL_MODBUS.Input_register_TCP_HMI[1030] := GVL_COM.COM_ADM100W_1.HMI_OUTPUT_L2_CURRENT.Word_value[0];                  // 1031 | ADM100W L2 Current (low word)
	GVL_MODBUS.Input_register_TCP_HMI[1031] := GVL_COM.COM_ADM100W_1.HMI_OUTPUT_L2_CURRENT.Word_value[1];                  // 1032 | ADM100W L2 Current (high word)
	GVL_MODBUS.Input_register_TCP_HMI[1032] := GVL_COM.COM_ADM100W_1.HMI_OUTPUT_L2_ACTIVE_POWER.Word_value[0];             // 1033 | ADM100W L2 Active Power (low word)
	GVL_MODBUS.Input_register_TCP_HMI[1033] := GVL_COM.COM_ADM100W_1.HMI_OUTPUT_L2_ACTIVE_POWER.Word_value[1];             // 1034 | ADM100W L2 Active Power (high word)
	GVL_MODBUS.Input_register_TCP_HMI[1034] := GVL_COM.COM_ADM100W_1.HMI_OUTPUT_L2_APPARENT_POWER.Word_value[0];           // 1035 | ADM100W L2 Apparent Power (low word)
	GVL_MODBUS.Input_register_TCP_HMI[1035] := GVL_COM.COM_ADM100W_1.HMI_OUTPUT_L2_APPARENT_POWER.Word_value[1];           // 1036 | ADM100W L2 Apparent Power (high word)
	GVL_MODBUS.Input_register_TCP_HMI[1036] := GVL_COM.COM_ADM100W_1.HMI_OUTPUT_L2_REACTIVE_POWER.Word_value[0];           // 1037 | ADM100W L2 Reactive Power (low word)
	GVL_MODBUS.Input_register_TCP_HMI[1037] := GVL_COM.COM_ADM100W_1.HMI_OUTPUT_L2_REACTIVE_POWER.Word_value[1];           // 1038 | ADM100W L2 Reactive Power (high word)
	GVL_MODBUS.Input_register_TCP_HMI[1038] := GVL_COM.COM_ADM100W_1.HMI_OUTPUT_L2_CURRENT_PHASE_ANGLE.Word_value[0];      // 1039 | ADM100W L2 Current Phase Angle (low word)
	GVL_MODBUS.Input_register_TCP_HMI[1039] := GVL_COM.COM_ADM100W_1.HMI_OUTPUT_L2_CURRENT_PHASE_ANGLE.Word_value[1];      // 1040 | ADM100W L2 Current Phase Angle (high word)
	GVL_MODBUS.Input_register_TCP_HMI[1040] := GVL_COM.COM_ADM100W_1.HMI_OUTPUT_L2_POWER_FACTOR.Word_value[0];             // 1041 | ADM100W L2 Power Factor (low word)
	GVL_MODBUS.Input_register_TCP_HMI[1041] := GVL_COM.COM_ADM100W_1.HMI_OUTPUT_L2_POWER_FACTOR.Word_value[1];             // 1042 | ADM100W L2 Power Factor (high word)
	GVL_MODBUS.Input_register_TCP_HMI[1042] := GVL_COM.COM_ADM100W_1.HMI_OUTPUT_L2_VOLTAGE_THD.Word_value[0];              // 1043 | ADM100W L2 Voltage THD (low word)
	GVL_MODBUS.Input_register_TCP_HMI[1043] := GVL_COM.COM_ADM100W_1.HMI_OUTPUT_L2_VOLTAGE_THD.Word_value[1];              // 1044 | ADM100W L2 Voltage THD (high word)
	GVL_MODBUS.Input_register_TCP_HMI[1044] := GVL_COM.COM_ADM100W_1.HMI_OUTPUT_L2_CURRENT_THD.Word_value[0];              // 1045 | ADM100W L2 Current THD (low word)
	GVL_MODBUS.Input_register_TCP_HMI[1045] := GVL_COM.COM_ADM100W_1.HMI_OUTPUT_L2_CURRENT_THD.Word_value[1];              // 1046 | ADM100W L2 Current THD (high word)
	GVL_MODBUS.Input_register_TCP_HMI[1046] := GVL_COM.COM_ADM100W_1.HMI_OUTPUT_L2_MAX_LOAD.Word_value[0];                 // 1047 | ADM100W L2 Max Load (low word)
	GVL_MODBUS.Input_register_TCP_HMI[1047] := GVL_COM.COM_ADM100W_1.HMI_OUTPUT_L2_MAX_LOAD.Word_value[1];                 // 1048 | ADM100W L2 Max Load (high word)
	GVL_MODBUS.Input_register_TCP_HMI[1048] := GVL_COM.COM_ADM100W_1.HMI_OUTPUT_L1_L3_VOLTAGE_PHASE_ANGLE.Word_value[0];   // 1049 | ADM100W L1-L3 Voltage Phase Angle (low word)
	GVL_MODBUS.Input_register_TCP_HMI[1049] := GVL_COM.COM_ADM100W_1.HMI_OUTPUT_L1_L3_VOLTAGE_PHASE_ANGLE.Word_value[1];   // 1050 | ADM100W L1-L3 Voltage Phase Angle (high word)
	GVL_MODBUS.Input_register_TCP_HMI[1050] := GVL_COM.COM_ADM100W_1.HMI_OUTPUT_L3_L1_VOLTAGE.Word_value[0];               // 1051 | ADM100W L3-L1 Voltage (low word)
	GVL_MODBUS.Input_register_TCP_HMI[1051] := GVL_COM.COM_ADM100W_1.HMI_OUTPUT_L3_L1_VOLTAGE.Word_value[1];               // 1052 | ADM100W L3-L1 Voltage (high word)
	GVL_MODBUS.Input_register_TCP_HMI[1052] := GVL_COM.COM_ADM100W_1.HMI_OUTPUT_L3_N_VOLTAGE.Word_value[0];                // 1053 | ADM100W L3-N Voltage (low word)
	GVL_MODBUS.Input_register_TCP_HMI[1053] := GVL_COM.COM_ADM100W_1.HMI_OUTPUT_L3_N_VOLTAGE.Word_value[1];                // 1054 | ADM100W L3-N Voltage (high word)
	GVL_MODBUS.Input_register_TCP_HMI[1054] := GVL_COM.COM_ADM100W_1.HMI_OUTPUT_L3_CURRENT.Word_value[0];                  // 1055 | ADM100W L3 Current (low word)
	GVL_MODBUS.Input_register_TCP_HMI[1055] := GVL_COM.COM_ADM100W_1.HMI_OUTPUT_L3_CURRENT.Word_value[1];                  // 1056 | ADM100W L3 Current (high word)
	GVL_MODBUS.Input_register_TCP_HMI[1056] := GVL_COM.COM_ADM100W_1.HMI_OUTPUT_L3_ACTIVE_POWER.Word_value[0];             // 1057 | ADM100W L3 Active Power (low word)
	GVL_MODBUS.Input_register_TCP_HMI[1057] := GVL_COM.COM_ADM100W_1.HMI_OUTPUT_L3_ACTIVE_POWER.Word_value[1];             // 1058 | ADM100W L3 Active Power (high word)
	GVL_MODBUS.Input_register_TCP_HMI[1058] := GVL_COM.COM_ADM100W_1.HMI_OUTPUT_L3_APPARENT_POWER.Word_value[0];           // 1059 | ADM100W L3 Apparent Power (low word)
	GVL_MODBUS.Input_register_TCP_HMI[1059] := GVL_COM.COM_ADM100W_1.HMI_OUTPUT_L3_APPARENT_POWER.Word_value[1];           // 1060 | ADM100W L3 Apparent Power (high word)
	GVL_MODBUS.Input_register_TCP_HMI[1060] := GVL_COM.COM_ADM100W_1.HMI_OUTPUT_L3_REACTIVE_POWER.Word_value[0];           // 1061 | ADM100W L3 Reactive Power (low word)
	GVL_MODBUS.Input_register_TCP_HMI[1061] := GVL_COM.COM_ADM100W_1.HMI_OUTPUT_L3_REACTIVE_POWER.Word_value[1];           // 1062 | ADM100W L3 Reactive Power (high word)
	GVL_MODBUS.Input_register_TCP_HMI[1062] := GVL_COM.COM_ADM100W_1.HMI_OUTPUT_L3_CURRENT_PHASE_ANGLE.Word_value[0];      // 1063 | ADM100W L3 Current Phase Angle (low word)
	GVL_MODBUS.Input_register_TCP_HMI[1063] := GVL_COM.COM_ADM100W_1.HMI_OUTPUT_L3_CURRENT_PHASE_ANGLE.Word_value[1];      // 1064 | ADM100W L3 Current Phase Angle (high word)
	GVL_MODBUS.Input_register_TCP_HMI[1064] := GVL_COM.COM_ADM100W_1.HMI_OUTPUT_L3_POWER_FACTOR.Word_value[0];             // 1065 | ADM100W L3 Power Factor (low word)
	GVL_MODBUS.Input_register_TCP_HMI[1065] := GVL_COM.COM_ADM100W_1.HMI_OUTPUT_L3_POWER_FACTOR.Word_value[1];             // 1066 | ADM100W L3 Power Factor (high word)
	GVL_MODBUS.Input_register_TCP_HMI[1066] := GVL_COM.COM_ADM100W_1.HMI_OUTPUT_L3_VOLTAGE_THD.Word_value[0];              // 1067 | ADM100W L3 Voltage THD (low word)
	GVL_MODBUS.Input_register_TCP_HMI[1067] := GVL_COM.COM_ADM100W_1.HMI_OUTPUT_L3_VOLTAGE_THD.Word_value[1];              // 1068 | ADM100W L3 Voltage THD (high word)
	GVL_MODBUS.Input_register_TCP_HMI[1068] := GVL_COM.COM_ADM100W_1.HMI_OUTPUT_L3_CURRENT_THD.Word_value[0];              // 1069 | ADM100W L3 Current THD (low word)
	GVL_MODBUS.Input_register_TCP_HMI[1069] := GVL_COM.COM_ADM100W_1.HMI_OUTPUT_L3_CURRENT_THD.Word_value[1];              // 1070 | ADM100W L3 Current THD (high word)
	GVL_MODBUS.Input_register_TCP_HMI[1070] := GVL_COM.COM_ADM100W_1.HMI_OUTPUT_L3_MAX_LOAD.Word_value[0];                 // 1071 | ADM100W L3 Max Load (low word)
	GVL_MODBUS.Input_register_TCP_HMI[1071] := GVL_COM.COM_ADM100W_1.HMI_OUTPUT_L3_MAX_LOAD.Word_value[1];                 // 1072 | ADM100W L3 Max Load (high word)
	GVL_MODBUS.Input_register_TCP_HMI[1072] := GVL_COM.COM_ADM100W_1.HMI_OUTPUT_INTERNAL_TEMPERATURE.Word_value[0];        // 1073 | ADM100W Internal Temperature (low word)
	GVL_MODBUS.Input_register_TCP_HMI[1073] := GVL_COM.COM_ADM100W_1.HMI_OUTPUT_INTERNAL_TEMPERATURE.Word_value[1];        // 1074 | ADM100W Internal Temperature (high word)
	GVL_MODBUS.Input_register_TCP_HMI[1074] := GVL_COM.COM_ADM100W_1.HMI_OUTPUT_ACTIVE_ENERGY.Word_value[0];               // 1075 | ADM100W Active Energy (low word)
	GVL_MODBUS.Input_register_TCP_HMI[1075] := GVL_COM.COM_ADM100W_1.HMI_OUTPUT_ACTIVE_ENERGY.Word_value[1];               // 1076 | ADM100W Active Energy (high word)
	GVL_MODBUS.Input_register_TCP_HMI[1076] := GVL_COM.COM_ADM100W_1.HMI_OUTPUT_APPARENT_ENERGY.Word_value[0];             // 1077 | ADM100W Apparent Energy (low word)
	GVL_MODBUS.Input_register_TCP_HMI[1077] := GVL_COM.COM_ADM100W_1.HMI_OUTPUT_APPARENT_ENERGY.Word_value[1];             // 1078 | ADM100W Apparent Energy (high word)
	GVL_MODBUS.Input_register_TCP_HMI[1078] := GVL_COM.COM_ADM100W_1.HMI_OUTPUT_REACTIVE_ENERGY.Word_value[0];             // 1079 | ADM100W Reactive Energy (low word)
	GVL_MODBUS.Input_register_TCP_HMI[1079] := GVL_COM.COM_ADM100W_1.HMI_OUTPUT_REACTIVE_ENERGY.Word_value[1];             // 1080 | ADM100W Reactive Energy (high word)
	GVL_MODBUS.Input_register_TCP_HMI[1080] := GVL_COM.COM_ADM100W_1.HMI_OUTPUT_TOTAL_ACTIVE_POWER.Word_value[0];          // 1081 | ADM100W Total Active Power (low word)
	GVL_MODBUS.Input_register_TCP_HMI[1081] := GVL_COM.COM_ADM100W_1.HMI_OUTPUT_TOTAL_ACTIVE_POWER.Word_value[1];          // 1082 | ADM100W Total Active Power (high word)
	GVL_MODBUS.Input_register_TCP_HMI[1082] := GVL_COM.COM_ADM100W_1.HMI_OUTPUT_TOTAL_APPARENT_POWER.Word_value[0];        // 1083 | ADM100W Total Apparent Power (low word)
	GVL_MODBUS.Input_register_TCP_HMI[1083] := GVL_COM.COM_ADM100W_1.HMI_OUTPUT_TOTAL_APPARENT_POWER.Word_value[1];        // 1084 | ADM100W Total Apparent Power (high word)
	GVL_MODBUS.Input_register_TCP_HMI[1084] := GVL_COM.COM_ADM100W_1.HMI_OUTPUT_TOTAL_REACTIVE_POWER.Word_value[0];        // 1085 | ADM100W Total Reactive Power (low word)
	GVL_MODBUS.Input_register_TCP_HMI[1085] := GVL_COM.COM_ADM100W_1.HMI_OUTPUT_TOTAL_REACTIVE_POWER.Word_value[1];        // 1086 | ADM100W Total Reactive Power (high word)
	GVL_MODBUS.Input_register_TCP_HMI[1086] := GVL_COM.COM_ADM100W_1.HMI_OUTPUT_ALL_PHASE_POWER_FACTOR.Word_value[0];      // 1087 | ADM100W All Phase Power Factor (low word)
	GVL_MODBUS.Input_register_TCP_HMI[1087] := GVL_COM.COM_ADM100W_1.HMI_OUTPUT_ALL_PHASE_POWER_FACTOR.Word_value[1];      // 1088 | ADM100W All Phase Power Factor (high word)

	//--- DOSENSOR_1
	GVL_MODBUS.Input_register_TCP_HMI[1088] := GVL_COM.COM_DOSENSOR_1.HMI_OUTPUT_SIGNAL.Word_value[0];   // 1089 | DO Sensor Signal (low word)
	GVL_MODBUS.Input_register_TCP_HMI[1089] := GVL_COM.COM_DOSENSOR_1.HMI_OUTPUT_SIGNAL.Word_value[1];   // 1090 | DO Sensor Signal (high word)

	//--- DIP1500_1
	GVL_MODBUS.Input_register_TCP_HMI[1090] := GVL_COM.COM_DIP1500_1.HMI_OUTPUT_FIRMWARE_VERSION;                               // 1091 | DIP1500 Firmware Version
	GVL_MODBUS.Input_register_TCP_HMI[1091] := GVL_COM.COM_DIP1500_1.HMI_OUTPUT_HARDWARE_VERSION;                               // 1092 | DIP1500 Hardware Version
	GVL_MODBUS.Input_register_TCP_HMI[1092] := GVL_COM.COM_DIP1500_1.HMI_OUTPUT_TEMPERATURE;                                    // 1093 | DIP1500 Temperature
	GVL_MODBUS.Input_register_TCP_HMI[1093] := GVL_COM.COM_DIP1500_1.HMI_OUTPUT_FLOAT_LEVEL_ALARM;                              // 1094 | DIP1500 Float Level Alarm
	GVL_MODBUS.Input_register_TCP_HMI[1094] := GVL_COM.COM_DIP1500_1.HMI_OUTPUT_DIGITAL_OUTPUT_VALUE;                           // 1095 | DIP1500 Digital Output Value
	GVL_MODBUS.Input_register_TCP_HMI[1095] := GVL_COM.COM_DIP1500_1.HMI_OUTPUT_REAL_TIME_RUN_TIME_OR_VOLUME.Word_value[0];     // 1096 | DIP1500 Real-Time Run Time Or Volume (low word)
	GVL_MODBUS.Input_register_TCP_HMI[1096] := GVL_COM.COM_DIP1500_1.HMI_OUTPUT_REAL_TIME_RUN_TIME_OR_VOLUME.Word_value[1];     // 1097 | DIP1500 Real-Time Run Time Or Volume (high word)
	GVL_MODBUS.Input_register_TCP_HMI[1097] := GVL_COM.COM_DIP1500_1.HMI_OUTPUT_ACCUMULATED_RUN_TIME_OR_VOLUME.Word_value[0];   // 1098 | DIP1500 Accumulated Run Time Or Volume (low word)
	GVL_MODBUS.Input_register_TCP_HMI[1098] := GVL_COM.COM_DIP1500_1.HMI_OUTPUT_ACCUMULATED_RUN_TIME_OR_VOLUME.Word_value[1];   // 1099 | DIP1500 Accumulated Run Time Or Volume (high word)

GFC_COM_OUT := TRUE;

                
END_FUNCTION

FUNCTION GFC_IO_IN : BOOL

                  
//==============================================================================
// GFC_IO_IN
// GVL_IOMAP (PLC I/O cards) -> GVL_IO
// Simple copies only, no conversion (conversions are done in the FBs)
//==============================================================================

//------------------------------------------------------------------------------
// Digital inputs
//------------------------------------------------------------------------------
	//--- DOSENSOR_1
	GVL_IO.IO_DOSENSOR_1.INPUT_SENSOR_FAULT := GVL_IOMAP.IOMAP_DI_FAULT_DOSENSOR_1;


//------------------------------------------------------------------------------
// Analog inputs
//------------------------------------------------------------------------------
	//--- DOSENSOR_1
	GVL_IO.IO_DOSENSOR_1.INPUT_SIGNAL := GVL_IOMAP.IOMAP_AI_SIGNAL_DOSENSOR_1;

GFC_IO_IN := TRUE;

                
END_FUNCTION

FUNCTION GFC_IO_OUT : BOOL

                  
//==============================================================================
// GFC_IO_OUT
// GVL_IO -> GVL_IOMAP (PLC I/O cards)
// Simple copies only, no conversion (conversions are done in the FBs)
//==============================================================================

//------------------------------------------------------------------------------
// Digital outputs
//------------------------------------------------------------------------------
	//--- DOSENSOR_1
	GVL_IOMAP.IOMAP_DO_HIGH_DOSENSOR_1 := GVL_IO.IO_DOSENSOR_1.OUTPUT_CALIBRATION_HIGH;
	GVL_IOMAP.IOMAP_DO_LOW_DOSENSOR_1  := GVL_IO.IO_DOSENSOR_1.OUTPUT_CALIBRATION_LOW;

GFC_IO_OUT := TRUE;

                
END_FUNCTION

FUNCTION_BLOCK FB_UPI_LOCAL_FUXA
  VAR_IN_OUT
    COM : DUT_COM_UPI_LOCAL_FUXA;  (* Requests and status with SCADA / HMI *)
    EXC : DUT_EXC_UPI_LOCAL_FUXA;  (* Status to equipment *)
  END_VAR
  VAR
    INTERN : DUT_INT_UPI_LOCAL_FUXA;  (* Internal variables *)
  END_VAR

                  
//==============================================================================
// FB_UPI_LOCAL_FUXA
// Global FUXA local mode for every equipment
// Set by the FUXA local request, reset by the FUXA auto request (pulse or maintained, auto wins)
// The equipment read this status through GFC_EXC_IN and report their own local status themselves
//==============================================================================

//------------------------------------------------------------------------------
// 1. INPUTS
//------------------------------------------------------------------------------
	INTERN.LOCAL_REQUEST := COM.SCADA_INPUT_LOCAL_REQUEST;
	INTERN.AUTO_REQUEST  := COM.SCADA_INPUT_AUTO_REQUEST;


//------------------------------------------------------------------------------
// 2. PROCESSING
//------------------------------------------------------------------------------
	IF INTERN.LOCAL_REQUEST THEN
		INTERN.LOCAL_ACTIVE := TRUE;
	END_IF
	IF INTERN.AUTO_REQUEST THEN
		INTERN.LOCAL_ACTIVE := FALSE;
	END_IF


//------------------------------------------------------------------------------
// 3. OUTPUTS
//------------------------------------------------------------------------------
	//--- EXC : to every equipment (through GFC_EXC_IN)
	EXC.UPI_OUTPUT_LOCAL_ACTIVE := INTERN.LOCAL_ACTIVE;

	//--- COM : status
	COM.SCADA_OUTPUT_LOCAL_ACTIVE := INTERN.LOCAL_ACTIVE;


                
END_FUNCTION_BLOCK

FUNCTION_BLOCK FB_UPI_LOCAL_HMI
  VAR_IN_OUT
    COM : DUT_COM_UPI_LOCAL_HMI;  (* Requests and status with SCADA / HMI *)
    EXC : DUT_EXC_UPI_LOCAL_HMI;  (* Status to equipment *)
  END_VAR
  VAR
    INTERN : DUT_INT_UPI_LOCAL_HMI;  (* Internal variables *)
  END_VAR

                  
//==============================================================================
// FB_UPI_LOCAL_HMI
// Global HMI local mode for every equipment
// Set by the HMI local request, reset by the HMI auto request (pulse or maintained, auto wins)
// The equipment read this status through GFC_EXC_IN and report their own local status themselves
//==============================================================================

//------------------------------------------------------------------------------
// 1. INPUTS
//------------------------------------------------------------------------------
	INTERN.LOCAL_REQUEST := COM.HMI_INPUT_LOCAL_REQUEST;
	INTERN.AUTO_REQUEST  := COM.HMI_INPUT_AUTO_REQUEST;


//------------------------------------------------------------------------------
// 2. PROCESSING
//------------------------------------------------------------------------------
	IF INTERN.LOCAL_REQUEST THEN
		INTERN.LOCAL_ACTIVE := TRUE;
	END_IF
	IF INTERN.AUTO_REQUEST THEN
		INTERN.LOCAL_ACTIVE := FALSE;
	END_IF


//------------------------------------------------------------------------------
// 3. OUTPUTS
//------------------------------------------------------------------------------
	//--- EXC : to every equipment (through GFC_EXC_IN)
	EXC.UPI_OUTPUT_LOCAL_ACTIVE := INTERN.LOCAL_ACTIVE;

	//--- COM : status
	COM.HMI_OUTPUT_LOCAL_ACTIVE   := INTERN.LOCAL_ACTIVE;
	COM.SCADA_OUTPUT_LOCAL_ACTIVE := INTERN.LOCAL_ACTIVE;   // also reported to FUXA


                
END_FUNCTION_BLOCK

FUNCTION_BLOCK GFB_INST
  VAR
    FB_ADM100W_1 : FB_INST_ADM100W;  (* Trumeter ADM100W power meter *)
    FB_DOSENSOR_1 : FB_INST_DOSENSOR;  (* Dissolved oxygen sensor *)
    FB_DIP1500_1 : FB_INST_DIP1500;  (* Kamoer DIP1500 peristaltic pump *)
  END_VAR

                  
//==============================================================================
// GFB_INST
// Calls every equipment instance
// One block per equipment, all interfaces connected
//==============================================================================

//--- ADM100W_1 : Trumeter ADM100W power meter
FB_ADM100W_1(
	PA  := GVL_PA.PA_ADM100W_1,
	COM := GVL_COM.COM_ADM100W_1,
	EXC := GVL_EXC.EXC_ADM100W_1,
	IO  := GVL_IO.IO_ADM100W_1);

//--- DOSENSOR_1 : Dissolved oxygen sensor
FB_DOSENSOR_1(
	PA  := GVL_PA.PA_DOSENSOR_1,
	COM := GVL_COM.COM_DOSENSOR_1,
	EXC := GVL_EXC.EXC_DOSENSOR_1,
	IO  := GVL_IO.IO_DOSENSOR_1);

//--- DIP1500_1 : Kamoer DIP1500 peristaltic pump
FB_DIP1500_1(
	PA  := GVL_PA.PA_DIP1500_1,
	COM := GVL_COM.COM_DIP1500_1,
	EXC := GVL_EXC.EXC_DIP1500_1,
	IO  := GVL_IO.IO_DIP1500_1);

                
END_FUNCTION_BLOCK

FUNCTION_BLOCK GFB_UPI
  VAR
    FB_UPI_LOCAL_FUXA_1 : FB_UPI_LOCAL_FUXA;  (* Global FUXA local mode *)
    FB_UPI_LOCAL_HMI_1 : FB_UPI_LOCAL_HMI;  (* Global HMI local mode *)
    FB_UPI_LOCAL_WEBVISU_1 : FB_UPI_LOCAL_WEBVISU;  (* Global WEBVISU local mode *)
  END_VAR

                  
//==============================================================================
// GFB_UPI
// Calls every functional unit (UPI)
// Runs before GFB_INST, results go to the equipment through GFC_EXC_IN
//==============================================================================

//--- UPI_LOCAL_FUXA : Global FUXA local mode
FB_UPI_LOCAL_FUXA_1(
	COM := GVL_COM.COM_UPI_LOCAL_FUXA,
	EXC := GVL_EXC.EXC_UPI_LOCAL_FUXA);

//--- UPI_LOCAL_HMI : Global HMI local mode
FB_UPI_LOCAL_HMI_1(
	COM := GVL_COM.COM_UPI_LOCAL_HMI,
	EXC := GVL_EXC.EXC_UPI_LOCAL_HMI);

//--- UPI_LOCAL_WEBVISU : Global WEBVISU local mode (direct IEC variables)
FB_UPI_LOCAL_WEBVISU_1(
	COM := GVL_COM.COM_UPI_LOCAL_WEBVISU,
	EXC := GVL_EXC.EXC_UPI_LOCAL_WEBVISU);

                
END_FUNCTION_BLOCK

FUNCTION_BLOCK FB_UPI_LOCAL_WEBVISU
  VAR_IN_OUT
    COM : DUT_COM_UPI_LOCAL_WEBVISU;  (* Direct IEC requests and status with WEBVISU *)
    EXC : DUT_EXC_UPI_LOCAL_WEBVISU;  (* Status to equipment *)
  END_VAR
  VAR
    INTERN : DUT_INT_UPI_LOCAL_WEBVISU;  (* Internal variables *)
  END_VAR

                  
//==============================================================================
// FB_UPI_LOCAL_WEBVISU
// Global WEBVISU local mode for every equipment
// Set by the WEBVISU local request, reset by the WEBVISU auto request (pulse or maintained, auto wins)
// The equipment read this status through GFC_EXC_IN and report their own local status themselves
//==============================================================================

//------------------------------------------------------------------------------
// 1. INPUTS
//------------------------------------------------------------------------------
	INTERN.LOCAL_REQUEST := COM.WEBVISU_INPUT_LOCAL_REQUEST;
	INTERN.AUTO_REQUEST  := COM.WEBVISU_INPUT_AUTO_REQUEST;


//------------------------------------------------------------------------------
// 2. PROCESSING
//------------------------------------------------------------------------------
	IF INTERN.LOCAL_REQUEST THEN
		INTERN.LOCAL_ACTIVE := TRUE;
	END_IF
	IF INTERN.AUTO_REQUEST THEN
		INTERN.LOCAL_ACTIVE := FALSE;
	END_IF


//------------------------------------------------------------------------------
// 3. OUTPUTS
//------------------------------------------------------------------------------
	//--- EXC : to every equipment (through GFC_EXC_IN)
	EXC.UPI_OUTPUT_LOCAL_ACTIVE := INTERN.LOCAL_ACTIVE;

	//--- COM : status
	COM.WEBVISU_OUTPUT_LOCAL_ACTIVE := INTERN.LOCAL_ACTIVE;


                
END_FUNCTION_BLOCK

FUNCTION FC_EXC_UPI_LOCAL_FUXA_ADM100W : BOOL
  VAR_IN_OUT
    EXC_UPI_LOCAL_FUXA : DUT_EXC_UPI_LOCAL_FUXA;  (* Exchanges of the UPI_LOCAL_FUXA instance *)
    EXC_ADM100W : DUT_EXC_ADM100W;  (* Exchanges of the ADM100W instance *)
  END_VAR

                  
//==============================================================================
// FC_EXC_UPI_LOCAL_FUXA_ADM100W
// Exchanges between one UPI_LOCAL_FUXA instance and one ADM100W instance
// Called in GFC_EXC, once per pair of instances, with their GVL_EXC variables
// Simple copies only, no conversion
//==============================================================================

//--- UPI_LOCAL_FUXA -> ADM100W
EXC_ADM100W.UPI_INPUT_GLOBAL_LOCAL_FUXA := EXC_UPI_LOCAL_FUXA.UPI_OUTPUT_LOCAL_ACTIVE;

FC_EXC_UPI_LOCAL_FUXA_ADM100W := TRUE;

                
END_FUNCTION

FUNCTION FC_EXC_UPI_LOCAL_FUXA_DIP1500 : BOOL
  VAR_IN_OUT
    EXC_UPI_LOCAL_FUXA : DUT_EXC_UPI_LOCAL_FUXA;  (* Exchanges of the UPI_LOCAL_FUXA instance *)
    EXC_DIP1500 : DUT_EXC_DIP1500;  (* Exchanges of the DIP1500 instance *)
  END_VAR

                  
//==============================================================================
// FC_EXC_UPI_LOCAL_FUXA_DIP1500
// Exchanges between one UPI_LOCAL_FUXA instance and one DIP1500 instance
// Called in GFC_EXC, once per pair of instances, with their GVL_EXC variables
// Simple copies only, no conversion
//==============================================================================

//--- UPI_LOCAL_FUXA -> DIP1500
EXC_DIP1500.UPI_INPUT_GLOBAL_LOCAL_FUXA := EXC_UPI_LOCAL_FUXA.UPI_OUTPUT_LOCAL_ACTIVE;

FC_EXC_UPI_LOCAL_FUXA_DIP1500 := TRUE;

                
END_FUNCTION

FUNCTION FC_EXC_UPI_LOCAL_FUXA_DOSENSOR : BOOL
  VAR_IN_OUT
    EXC_UPI_LOCAL_FUXA : DUT_EXC_UPI_LOCAL_FUXA;  (* Exchanges of the UPI_LOCAL_FUXA instance *)
    EXC_DOSENSOR : DUT_EXC_DOSENSOR;  (* Exchanges of the DOSENSOR instance *)
  END_VAR

                  
//==============================================================================
// FC_EXC_UPI_LOCAL_FUXA_DOSENSOR
// Exchanges between one UPI_LOCAL_FUXA instance and one DOSENSOR instance
// Called in GFC_EXC, once per pair of instances, with their GVL_EXC variables
// Simple copies only, no conversion
//==============================================================================

//--- UPI_LOCAL_FUXA -> DOSENSOR
EXC_DOSENSOR.UPI_INPUT_GLOBAL_LOCAL_FUXA := EXC_UPI_LOCAL_FUXA.UPI_OUTPUT_LOCAL_ACTIVE;

FC_EXC_UPI_LOCAL_FUXA_DOSENSOR := TRUE;

                
END_FUNCTION

FUNCTION FC_EXC_UPI_LOCAL_HMI_ADM100W : BOOL
  VAR_IN_OUT
    EXC_UPI_LOCAL_HMI : DUT_EXC_UPI_LOCAL_HMI;  (* Exchanges of the UPI_LOCAL_HMI instance *)
    EXC_ADM100W : DUT_EXC_ADM100W;  (* Exchanges of the ADM100W instance *)
  END_VAR

                  
//==============================================================================
// FC_EXC_UPI_LOCAL_HMI_ADM100W
// Exchanges between one UPI_LOCAL_HMI instance and one ADM100W instance
// Called in GFC_EXC, once per pair of instances, with their GVL_EXC variables
// Simple copies only, no conversion
//==============================================================================

//--- UPI_LOCAL_HMI -> ADM100W
EXC_ADM100W.UPI_INPUT_GLOBAL_LOCAL_HMI := EXC_UPI_LOCAL_HMI.UPI_OUTPUT_LOCAL_ACTIVE;

FC_EXC_UPI_LOCAL_HMI_ADM100W := TRUE;

                
END_FUNCTION

FUNCTION FC_EXC_UPI_LOCAL_HMI_DIP1500 : BOOL
  VAR_IN_OUT
    EXC_UPI_LOCAL_HMI : DUT_EXC_UPI_LOCAL_HMI;  (* Exchanges of the UPI_LOCAL_HMI instance *)
    EXC_DIP1500 : DUT_EXC_DIP1500;  (* Exchanges of the DIP1500 instance *)
  END_VAR

                  
//==============================================================================
// FC_EXC_UPI_LOCAL_HMI_DIP1500
// Exchanges between one UPI_LOCAL_HMI instance and one DIP1500 instance
// Called in GFC_EXC, once per pair of instances, with their GVL_EXC variables
// Simple copies only, no conversion
//==============================================================================

//--- UPI_LOCAL_HMI -> DIP1500
EXC_DIP1500.UPI_INPUT_GLOBAL_LOCAL_HMI := EXC_UPI_LOCAL_HMI.UPI_OUTPUT_LOCAL_ACTIVE;

FC_EXC_UPI_LOCAL_HMI_DIP1500 := TRUE;

                
END_FUNCTION

FUNCTION FC_EXC_UPI_LOCAL_HMI_DOSENSOR : BOOL
  VAR_IN_OUT
    EXC_UPI_LOCAL_HMI : DUT_EXC_UPI_LOCAL_HMI;  (* Exchanges of the UPI_LOCAL_HMI instance *)
    EXC_DOSENSOR : DUT_EXC_DOSENSOR;  (* Exchanges of the DOSENSOR instance *)
  END_VAR

                  
//==============================================================================
// FC_EXC_UPI_LOCAL_HMI_DOSENSOR
// Exchanges between one UPI_LOCAL_HMI instance and one DOSENSOR instance
// Called in GFC_EXC, once per pair of instances, with their GVL_EXC variables
// Simple copies only, no conversion
//==============================================================================

//--- UPI_LOCAL_HMI -> DOSENSOR
EXC_DOSENSOR.UPI_INPUT_GLOBAL_LOCAL_HMI := EXC_UPI_LOCAL_HMI.UPI_OUTPUT_LOCAL_ACTIVE;

FC_EXC_UPI_LOCAL_HMI_DOSENSOR := TRUE;

                
END_FUNCTION

FUNCTION FC_EXC_UPI_LOCAL_WEBVISU_ADM100W : BOOL
  VAR_IN_OUT
    EXC_UPI_LOCAL_WEBVISU : DUT_EXC_UPI_LOCAL_WEBVISU;  (* Exchanges of the UPI_LOCAL_WEBVISU instance *)
    EXC_ADM100W : DUT_EXC_ADM100W;  (* Exchanges of the ADM100W instance *)
  END_VAR

                  
//==============================================================================
// FC_EXC_UPI_LOCAL_WEBVISU_ADM100W
// Exchanges between one UPI_LOCAL_WEBVISU instance and one ADM100W instance
// Called in GFC_EXC, once per pair of instances, with their GVL_EXC variables
// Simple copies only, no conversion
//==============================================================================

//--- UPI_LOCAL_WEBVISU -> ADM100W
EXC_ADM100W.UPI_INPUT_GLOBAL_LOCAL_WEBVISU := EXC_UPI_LOCAL_WEBVISU.UPI_OUTPUT_LOCAL_ACTIVE;

FC_EXC_UPI_LOCAL_WEBVISU_ADM100W := TRUE;

                
END_FUNCTION

FUNCTION FC_EXC_UPI_LOCAL_WEBVISU_DIP1500 : BOOL
  VAR_IN_OUT
    EXC_UPI_LOCAL_WEBVISU : DUT_EXC_UPI_LOCAL_WEBVISU;  (* Exchanges of the UPI_LOCAL_WEBVISU instance *)
    EXC_DIP1500 : DUT_EXC_DIP1500;  (* Exchanges of the DIP1500 instance *)
  END_VAR

                  
//==============================================================================
// FC_EXC_UPI_LOCAL_WEBVISU_DIP1500
// Exchanges between one UPI_LOCAL_WEBVISU instance and one DIP1500 instance
// Called in GFC_EXC, once per pair of instances, with their GVL_EXC variables
// Simple copies only, no conversion
//==============================================================================

//--- UPI_LOCAL_WEBVISU -> DIP1500
EXC_DIP1500.UPI_INPUT_GLOBAL_LOCAL_WEBVISU := EXC_UPI_LOCAL_WEBVISU.UPI_OUTPUT_LOCAL_ACTIVE;

FC_EXC_UPI_LOCAL_WEBVISU_DIP1500 := TRUE;

                
END_FUNCTION

FUNCTION FC_EXC_UPI_LOCAL_WEBVISU_DOSENSOR : BOOL
  VAR_IN_OUT
    EXC_UPI_LOCAL_WEBVISU : DUT_EXC_UPI_LOCAL_WEBVISU;  (* Exchanges of the UPI_LOCAL_WEBVISU instance *)
    EXC_DOSENSOR : DUT_EXC_DOSENSOR;  (* Exchanges of the DOSENSOR instance *)
  END_VAR

                  
//==============================================================================
// FC_EXC_UPI_LOCAL_WEBVISU_DOSENSOR
// Exchanges between one UPI_LOCAL_WEBVISU instance and one DOSENSOR instance
// Called in GFC_EXC, once per pair of instances, with their GVL_EXC variables
// Simple copies only, no conversion
//==============================================================================

//--- UPI_LOCAL_WEBVISU -> DOSENSOR
EXC_DOSENSOR.UPI_INPUT_GLOBAL_LOCAL_WEBVISU := EXC_UPI_LOCAL_WEBVISU.UPI_OUTPUT_LOCAL_ACTIVE;

FC_EXC_UPI_LOCAL_WEBVISU_DOSENSOR := TRUE;

                
END_FUNCTION

FUNCTION GFC_EXC : BOOL

                  
//==============================================================================
// GFC_EXC
// Exchanges between instances : one FC_EXC_<A>_<B> call per pair of instances
// Called after GFB_UPI and before GFB_INST
//==============================================================================

//------------------------------------------------------------------------------
// ADM100W_1
//------------------------------------------------------------------------------
	//--- UPI_LOCAL_FUXA <-> ADM100W_1
	FC_EXC_UPI_LOCAL_FUXA_ADM100W(
		EXC_UPI_LOCAL_FUXA := GVL_EXC.EXC_UPI_LOCAL_FUXA,
		EXC_ADM100W        := GVL_EXC.EXC_ADM100W_1);

	//--- UPI_LOCAL_HMI <-> ADM100W_1
	FC_EXC_UPI_LOCAL_HMI_ADM100W(
		EXC_UPI_LOCAL_HMI := GVL_EXC.EXC_UPI_LOCAL_HMI,
		EXC_ADM100W       := GVL_EXC.EXC_ADM100W_1);

	//--- UPI_LOCAL_WEBVISU <-> ADM100W_1
	FC_EXC_UPI_LOCAL_WEBVISU_ADM100W(
		EXC_UPI_LOCAL_WEBVISU := GVL_EXC.EXC_UPI_LOCAL_WEBVISU,
		EXC_ADM100W           := GVL_EXC.EXC_ADM100W_1);


//------------------------------------------------------------------------------
// DOSENSOR_1
//------------------------------------------------------------------------------
	//--- UPI_LOCAL_FUXA <-> DOSENSOR_1
	FC_EXC_UPI_LOCAL_FUXA_DOSENSOR(
		EXC_UPI_LOCAL_FUXA := GVL_EXC.EXC_UPI_LOCAL_FUXA,
		EXC_DOSENSOR       := GVL_EXC.EXC_DOSENSOR_1);

	//--- UPI_LOCAL_HMI <-> DOSENSOR_1
	FC_EXC_UPI_LOCAL_HMI_DOSENSOR(
		EXC_UPI_LOCAL_HMI := GVL_EXC.EXC_UPI_LOCAL_HMI,
		EXC_DOSENSOR      := GVL_EXC.EXC_DOSENSOR_1);

	//--- UPI_LOCAL_WEBVISU <-> DOSENSOR_1
	FC_EXC_UPI_LOCAL_WEBVISU_DOSENSOR(
		EXC_UPI_LOCAL_WEBVISU := GVL_EXC.EXC_UPI_LOCAL_WEBVISU,
		EXC_DOSENSOR          := GVL_EXC.EXC_DOSENSOR_1);


//------------------------------------------------------------------------------
// DIP1500_1
//------------------------------------------------------------------------------
	//--- UPI_LOCAL_FUXA <-> DIP1500_1
	FC_EXC_UPI_LOCAL_FUXA_DIP1500(
		EXC_UPI_LOCAL_FUXA := GVL_EXC.EXC_UPI_LOCAL_FUXA,
		EXC_DIP1500        := GVL_EXC.EXC_DIP1500_1);

	//--- UPI_LOCAL_HMI <-> DIP1500_1
	FC_EXC_UPI_LOCAL_HMI_DIP1500(
		EXC_UPI_LOCAL_HMI := GVL_EXC.EXC_UPI_LOCAL_HMI,
		EXC_DIP1500       := GVL_EXC.EXC_DIP1500_1);

	//--- UPI_LOCAL_WEBVISU <-> DIP1500_1
	FC_EXC_UPI_LOCAL_WEBVISU_DIP1500(
		EXC_UPI_LOCAL_WEBVISU := GVL_EXC.EXC_UPI_LOCAL_WEBVISU,
		EXC_DIP1500           := GVL_EXC.EXC_DIP1500_1);

GFC_EXC := TRUE;

                
END_FUNCTION

PROGRAM PLC_PRG
  VAR
    GFB_UPI_1 : GFB_UPI;  (* Functional units *)
    GFB_INST_1 : GFB_INST;  (* Equipment instances *)
  END_VAR

                  
//==============================================================================
// PLC_PRG
// Main cycle : 1. read all inputs, 2. functional units, 3. equipment, 4. write all outputs
//==============================================================================

//------------------------------------------------------------------------------
// 1. INPUTS : interfaces -> GVL
//------------------------------------------------------------------------------
GFC_COM_IN();
GFC_IO_IN();

//------------------------------------------------------------------------------
// 2. FUNCTIONAL UNITS (UPI) and exchanges between instances
//------------------------------------------------------------------------------
GFB_UPI_1();
GFC_EXC();      // exchanges between instances (FC_EXC_...)

//------------------------------------------------------------------------------
// 3. EQUIPMENT
//------------------------------------------------------------------------------
GFB_INST_1();

//------------------------------------------------------------------------------
// 4. OUTPUTS : GVL -> interfaces
//------------------------------------------------------------------------------
GFC_COM_OUT();
GFC_IO_OUT();

                
END_PROGRAM

CONFIGURATION Application
  RESOURCE Application ON PLC
    VAR_GLOBAL  (* GVL_MODBUS *)
      Coils_TCP_HMI : ARRAY[0..187] OF BYTE;  (* -----------------Modbus TCP line IHM -> API (coils, %IX) *)
      Discret_input_TCP_HMI : ARRAY[0..187] OF BYTE;  (* API -> IHM (entrées discrètes, %QX) *)
      Holding_register_TCP_HMI : ARRAY[0..1500] OF WORD;  (* IHM -> API (registres de retenue, %IW) *)
      Input_register_TCP_HMI : ARRAY[0..1500] OF WORD;  (* API -> IHM (registres d'entrée, %QW) *)
      ADM100W_InputRegisters : ARRAY[0..87] OF WORD;  (* ------------------Modbus RTU line ---ADM100W *)
      ADM100W_Alarms : ARRAY[0..1] OF BYTE;
      DIP1500_Coils : ARRAY[0..3] OF BOOL;  (* ---Kamoer DIP1500 Coils - wrinting to pump *)
      DIP1500_InputRegisters : ARRAY[0..4] OF WORD;  (* input register - reading from pump *)
      DIP1500_Holding_Cmd : ARRAY[0..5] OF WORD;  (* Discrete input Holding registers - Writing to pump *)
      DIP1500_Holding_Config : ARRAY[0..6] OF WORD;
      DIP1500_Holding_Counters : ARRAY[0..3] OF WORD;  (* Holding registers - Reading from pump *)
    END_VAR
    {attribute 'qualified_only'}
    VAR_GLOBAL  (* GVL_IO *)
      IO_ADM100W_1 : DUT_IO_ADM100W;  (* Trumeter ADM100W power meter *)
      IO_DOSENSOR_1 : DUT_IO_DOSENSOR;  (* Dissolved oxygen sensor *)
      IO_DIP1500_1 : DUT_IO_DIP1500;  (* Kamoer DIP1500 peristaltic pump *)
    END_VAR
    {attribute 'qualified_only'}
    VAR_GLOBAL  (* GVL_IOMAP *)
      IOMAP_AI_SIGNAL_DOSENSOR_1 : DWORD;
      IOMAP_DI_FAULT_DOSENSOR_1 : BOOL;
      IOMAP_DO_HIGH_DOSENSOR_1 : BOOL;
      IOMAP_DO_LOW_DOSENSOR_1 : BOOL;
    END_VAR
    {attribute 'qualified_only'}
    VAR_GLOBAL  (* GVL_COM *)
      COM_ADM100W_1 : DUT_COM_ADM100W;  (* Trumeter ADM100W power meter *)
      COM_DOSENSOR_1 : DUT_COM_DOSENSOR;  (* Dissolved oxygen sensor *)
      COM_DIP1500_1 : DUT_COM_DIP1500;  (* Kamoer DIP1500 peristaltic pump *)
      COM_UPI_LOCAL_FUXA : DUT_COM_UPI_LOCAL_FUXA;  (* Global FUXA local mode *)
      COM_UPI_LOCAL_HMI : DUT_COM_UPI_LOCAL_HMI;  (* Global HMI local mode *)
      COM_UPI_LOCAL_WEBVISU : DUT_COM_UPI_LOCAL_WEBVISU;  (* Global WEBVISU local mode *)
    END_VAR
    {attribute 'qualified_only'}
    VAR_GLOBAL  (* GVL_EXC *)
      EXC_ADM100W_1 : DUT_EXC_ADM100W;  (* Trumeter ADM100W power meter *)
      EXC_DOSENSOR_1 : DUT_EXC_DOSENSOR;  (* Dissolved oxygen sensor *)
      EXC_DIP1500_1 : DUT_EXC_DIP1500;  (* Kamoer DIP1500 peristaltic pump *)
      EXC_UPI_LOCAL_FUXA : DUT_EXC_UPI_LOCAL_FUXA;  (* Global FUXA local mode *)
      EXC_UPI_LOCAL_HMI : DUT_EXC_UPI_LOCAL_HMI;  (* Global HMI local mode *)
      EXC_UPI_LOCAL_WEBVISU : DUT_EXC_UPI_LOCAL_WEBVISU;  (* Global WEBVISU local mode *)
    END_VAR
    {attribute 'qualified_only'}
    {attribute 'checksumnoinit_override' := '3446479488'}
    {attribute 'init_related_code' := '6eea8fa9-da21-468e-bab1-ddc04c20a5e9'}
    VAR_GLOBAL RETAIN PERSISTENT  (* GVL_PA *)
      {attribute 'order_in_persistent_editor' := '0'}
      PA_ADM100W_1 : DUT_PA_ADM100W;  (* Trumeter ADM100W power meter *)
      {attribute 'order_in_persistent_editor' := '1'}
      PA_DOSENSOR_1 : DUT_PA_DOSENSOR;  (* Dissolved oxygen sensor *)
      {attribute 'order_in_persistent_editor' := '2'}
      PA_DIP1500_1 : DUT_PA_DIP1500;  (* Kamoer DIP1500 peristaltic pump *)
    END_VAR
  END_RESOURCE
END_CONFIGURATION
